FUNCTION_BLOCK FB_Counter
VAR_INPUT
    enable : BOOL;
END_VAR
VAR_OUTPUT
    count : DINT;
END_VAR

IF enable THEN
    count := count + 1;
END_IF;

END_FUNCTION_BLOCK

(* stored: Version 1.1.0.1, ProductVersion 3.1.4026.0
   POU FB_Counter: Id {0342b13c-6f0c-4a32-a6b9-44604cf44317} *)
